// LS Electric XG5000 project: elb
// PLC LSPLC
// module base 0 slot 0: 입출력 모듈:XBC-DR32H (DC 24V 입력, 릴레이 출력 32점)
// module base 0 slot 1: 입력 모듈:XBE-DC16A/B (DC24V 입력, 16점 / DC12/24V 입력, 16점)

PROGRAM 스위치_입력 (task: 스캔 프로그램)

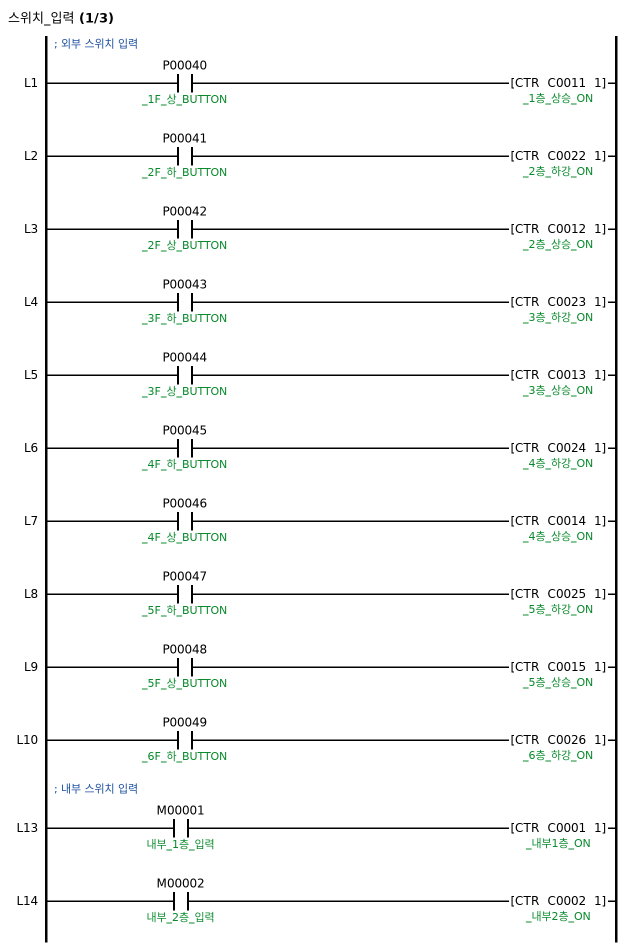
// 외부 스위치 입력
; L1
LOAD      P00040	// _1F_상_BUTTON
CTR       C0011 1	// _1층_상승_ON
; L2
LOAD      P00041	// _2F_하_BUTTON
CTR       C0022 1	// _2층_하강_ON
; L3
LOAD      P00042	// _2F_상_BUTTON
CTR       C0012 1	// _2층_상승_ON
; L4
LOAD      P00043	// _3F_하_BUTTON
CTR       C0023 1	// _3층_하강_ON
; L5
LOAD      P00044	// _3F_상_BUTTON
CTR       C0013 1	// _3층_상승_ON
; L6
LOAD      P00045	// _4F_하_BUTTON
CTR       C0024 1	// _4층_하강_ON
; L7
LOAD      P00046	// _4F_상_BUTTON
CTR       C0014 1	// _4층_상승_ON
; L8
LOAD      P00047	// _5F_하_BUTTON
CTR       C0025 1	// _5층_하강_ON
; L9
LOAD      P00048	// _5F_상_BUTTON
CTR       C0015 1	// _5층_상승_ON
; L10
LOAD      P00049	// _6F_하_BUTTON
CTR       C0026 1	// _6층_하강_ON
// 내부 스위치 입력
; L13
LOAD      M00001	// 내부_1층_입력
CTR       C0001 1	// _내부1층_ON
; L14
LOAD      M00002	// 내부_2층_입력
CTR       C0002 1	// _내부2층_ON

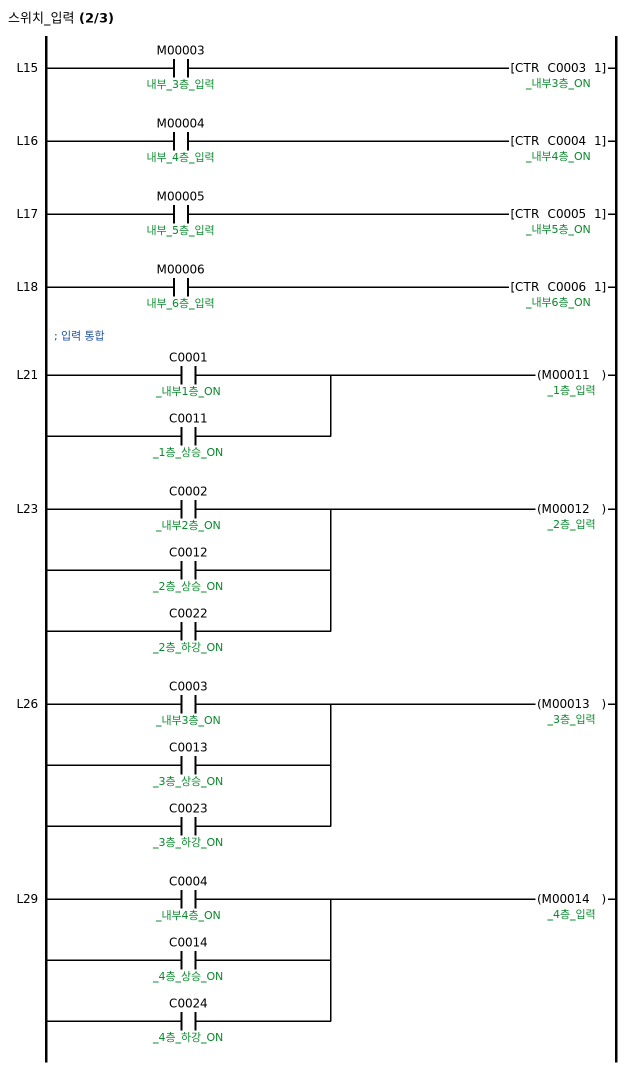
; L15
LOAD      M00003	// 내부_3층_입력
CTR       C0003 1	// _내부3층_ON
; L16
LOAD      M00004	// 내부_4층_입력
CTR       C0004 1	// _내부4층_ON
; L17
LOAD      M00005	// 내부_5층_입력
CTR       C0005 1	// _내부5층_ON
; L18
LOAD      M00006	// 내부_6층_입력
CTR       C0006 1	// _내부6층_ON
// 입력 통합
; L21
LOAD      C0001	// _내부1층_ON
OR        C0011	// _1층_상승_ON
OUT       M00011	// _1층_입력
; L23
LOAD      C0002	// _내부2층_ON
OR        C0012	// _2층_상승_ON
OR        C0022	// _2층_하강_ON
OUT       M00012	// _2층_입력
; L26
LOAD      C0003	// _내부3층_ON
OR        C0013	// _3층_상승_ON
OR        C0023	// _3층_하강_ON
OUT       M00013	// _3층_입력
; L29
LOAD      C0004	// _내부4층_ON
OR        C0014	// _4층_상승_ON
OR        C0024	// _4층_하강_ON
OUT       M00014	// _4층_입력

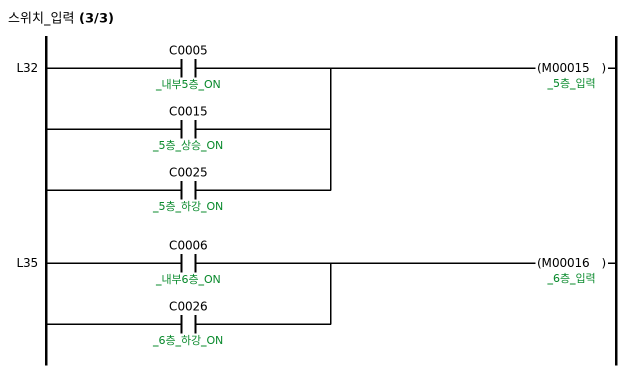
; L32
LOAD      C0005	// _내부5층_ON
OR        C0015	// _5층_상승_ON
OR        C0025	// _5층_하강_ON
OUT       M00015	// _5층_입력
; L35
LOAD      C0006	// _내부6층_ON
OR        C0026	// _6층_하강_ON
OUT       M00016	// _6층_입력

PROGRAM 센서감지(현재위치 (task: 스캔 프로그램)

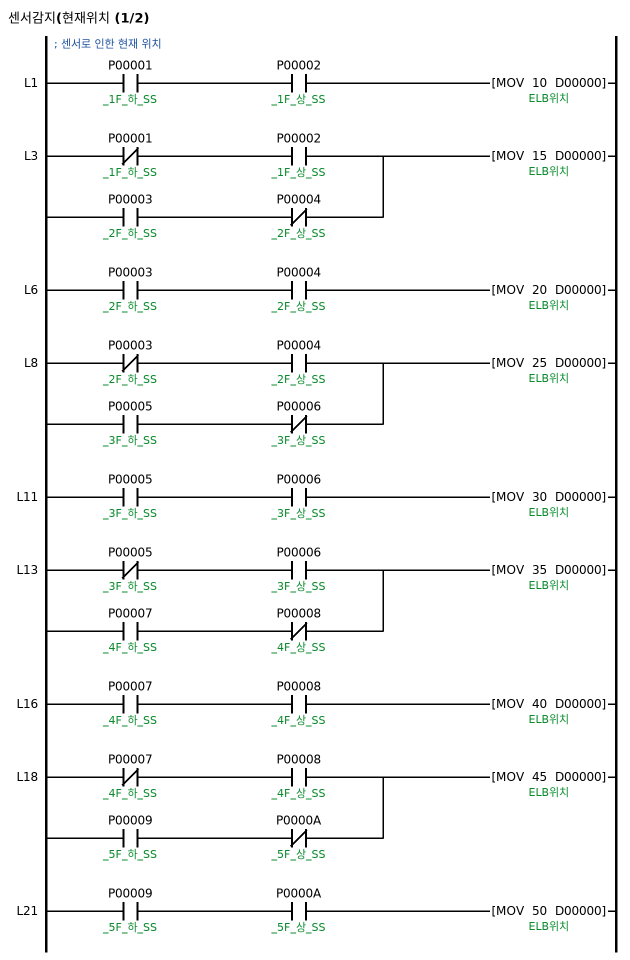
// 센서로 인한 현재 위치
; L1
LOAD      P00001	// _1F_하_SS
AND       P00002	// _1F_상_SS
MOV       10 D00000	// ELB위치
; L3
LOAD NOT  P00001	// _1F_하_SS
AND       P00002	// _1F_상_SS
LOAD      P00003	// _2F_하_SS
AND NOT   P00004	// _2F_상_SS
OR LOAD
MOV       15 D00000	// ELB위치
; L6
LOAD      P00003	// _2F_하_SS
AND       P00004	// _2F_상_SS
MOV       20 D00000	// ELB위치
; L8
LOAD NOT  P00003	// _2F_하_SS
AND       P00004	// _2F_상_SS
LOAD      P00005	// _3F_하_SS
AND NOT   P00006	// _3F_상_SS
OR LOAD
MOV       25 D00000	// ELB위치
; L11
LOAD      P00005	// _3F_하_SS
AND       P00006	// _3F_상_SS
MOV       30 D00000	// ELB위치
; L13
LOAD NOT  P00005	// _3F_하_SS
AND       P00006	// _3F_상_SS
LOAD      P00007	// _4F_하_SS
AND NOT   P00008	// _4F_상_SS
OR LOAD
MOV       35 D00000	// ELB위치
; L16
LOAD      P00007	// _4F_하_SS
AND       P00008	// _4F_상_SS
MOV       40 D00000	// ELB위치
; L18
LOAD NOT  P00007	// _4F_하_SS
AND       P00008	// _4F_상_SS
LOAD      P00009	// _5F_하_SS
AND NOT   P0000A	// _5F_상_SS
OR LOAD
MOV       45 D00000	// ELB위치
; L21
LOAD      P00009	// _5F_하_SS
AND       P0000A	// _5F_상_SS
MOV       50 D00000	// ELB위치

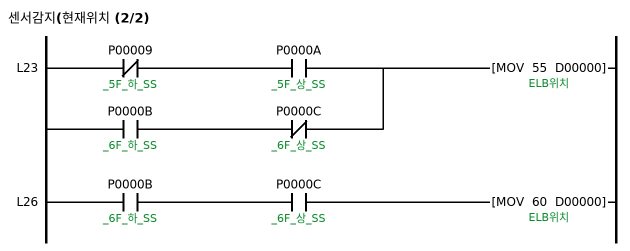
; L23
LOAD NOT  P00009	// _5F_하_SS
AND       P0000A	// _5F_상_SS
LOAD      P0000B	// _6F_하_SS
AND NOT   P0000C	// _6F_상_SS
OR LOAD
MOV       55 D00000	// ELB위치
; L26
LOAD      P0000B	// _6F_하_SS
AND       P0000C	// _6F_상_SS
MOV       60 D00000	// ELB위치

PROGRAM 모드전환 (task: 스캔 프로그램)

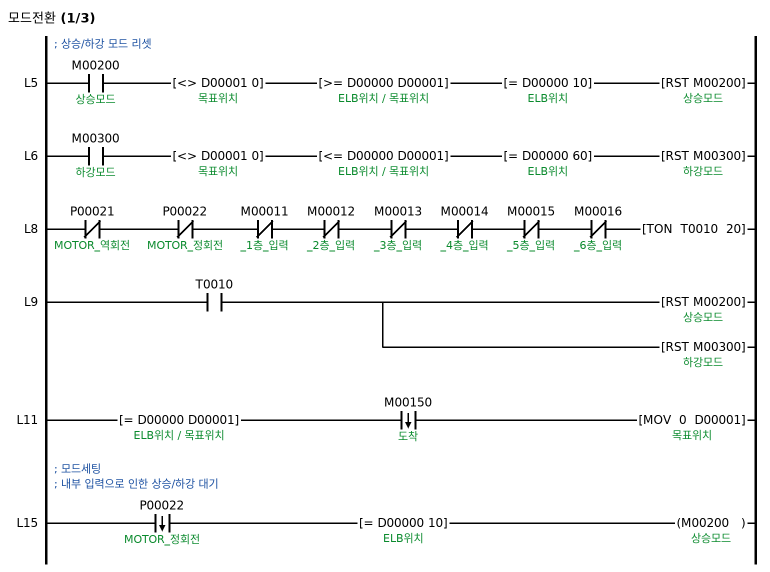
// 상승/하강 모드 리셋
; L5
LOAD      M00200	// 상승모드
AND<>     D00001 0	// 목표위치
AND>=     D00000 D00001	// ELB위치 / 목표위치
AND=      D00000 10	// ELB위치
RST       M00200	// 상승모드
; L6
LOAD      M00300	// 하강모드
AND<>     D00001 0	// 목표위치
AND<=     D00000 D00001	// ELB위치 / 목표위치
AND=      D00000 60	// ELB위치
RST       M00300	// 하강모드
; L8
LOAD NOT  P00021	// MOTOR_역회전
AND NOT   P00022	// MOTOR_정회전
AND NOT   M00011	// _1층_입력
AND NOT   M00012	// _2층_입력
AND NOT   M00013	// _3층_입력
AND NOT   M00014	// _4층_입력
AND NOT   M00015	// _5층_입력
AND NOT   M00016	// _6층_입력
TON       T0010 20
; L9
LOAD      T0010
RST       M00200	// 상승모드
RST       M00300	// 하강모드
; L11
LOAD=     D00000 D00001	// ELB위치 / 목표위치
ANDN      M00150	// 도착
MOV       0 D00001	// 목표위치
// 모드세팅
// 내부 입력으로 인한 상승/하강 대기
; L15
LOADN     P00022	// MOTOR_정회전
AND=      D00000 10	// ELB위치
OUT       M00200	// 상승모드

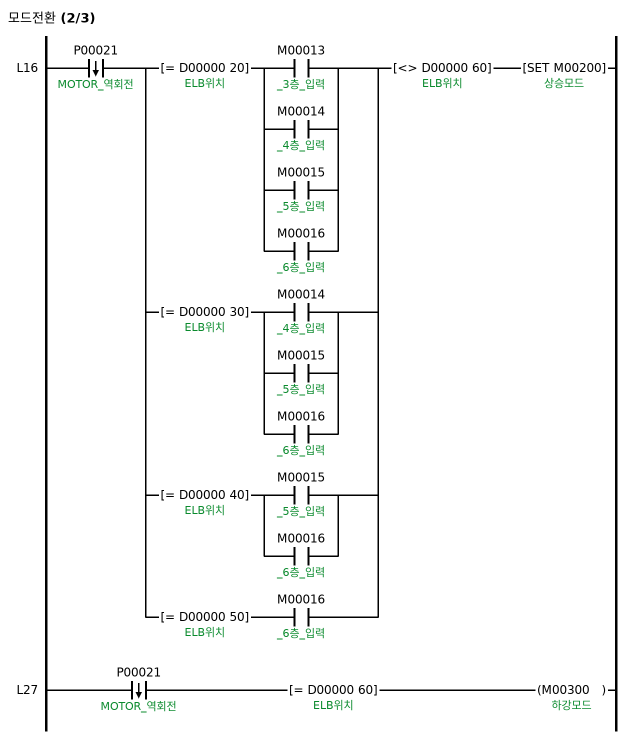
; L16
LOADN     P00021	// MOTOR_역회전
LOAD=     D00000 20	// ELB위치
LOAD      M00013	// _3층_입력
OR        M00014	// _4층_입력
OR        M00015	// _5층_입력
OR        M00016	// _6층_입력
AND LOAD
LOAD=     D00000 30	// ELB위치
LOAD      M00014	// _4층_입력
OR        M00015	// _5층_입력
OR        M00016	// _6층_입력
AND LOAD
OR LOAD
LOAD=     D00000 40	// ELB위치
LOAD      M00015	// _5층_입력
OR        M00016	// _6층_입력
AND LOAD
OR LOAD
LOAD=     D00000 50	// ELB위치
AND       M00016	// _6층_입력
OR LOAD
AND LOAD
AND<>     D00000 60	// ELB위치
SET       M00200	// 상승모드
; L27
LOADN     P00021	// MOTOR_역회전
AND=      D00000 60	// ELB위치
OUT       M00300	// 하강모드

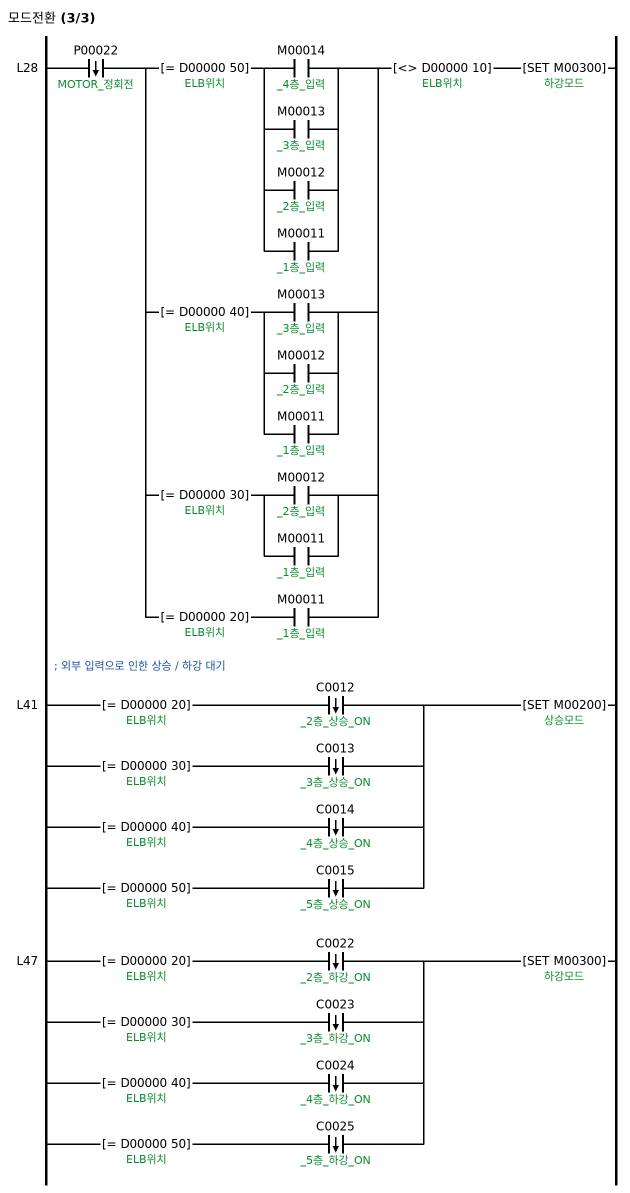
; L28
LOADN     P00022	// MOTOR_정회전
LOAD=     D00000 50	// ELB위치
LOAD      M00014	// _4층_입력
OR        M00013	// _3층_입력
OR        M00012	// _2층_입력
OR        M00011	// _1층_입력
AND LOAD
LOAD=     D00000 40	// ELB위치
LOAD      M00013	// _3층_입력
OR        M00012	// _2층_입력
OR        M00011	// _1층_입력
AND LOAD
OR LOAD
LOAD=     D00000 30	// ELB위치
LOAD      M00012	// _2층_입력
OR        M00011	// _1층_입력
AND LOAD
OR LOAD
LOAD=     D00000 20	// ELB위치
AND       M00011	// _1층_입력
OR LOAD
AND LOAD
AND<>     D00000 10	// ELB위치
SET       M00300	// 하강모드
// 외부 입력으로 인한 상승 / 하강 대기
; L41
LOAD=     D00000 20	// ELB위치
ANDN      C0012	// _2층_상승_ON
LOAD=     D00000 30	// ELB위치
ANDN      C0013	// _3층_상승_ON
OR LOAD
LOAD=     D00000 40	// ELB위치
ANDN      C0014	// _4층_상승_ON
OR LOAD
LOAD=     D00000 50	// ELB위치
ANDN      C0015	// _5층_상승_ON
OR LOAD
SET       M00200	// 상승모드
; L47
LOAD=     D00000 20	// ELB위치
ANDN      C0022	// _2층_하강_ON
LOAD=     D00000 30	// ELB위치
ANDN      C0023	// _3층_하강_ON
OR LOAD
LOAD=     D00000 40	// ELB위치
ANDN      C0024	// _4층_하강_ON
OR LOAD
LOAD=     D00000 50	// ELB위치
ANDN      C0025	// _5층_하강_ON
OR LOAD
SET       M00300	// 하강모드

PROGRAM 스위치리셋 (task: 스캔 프로그램)

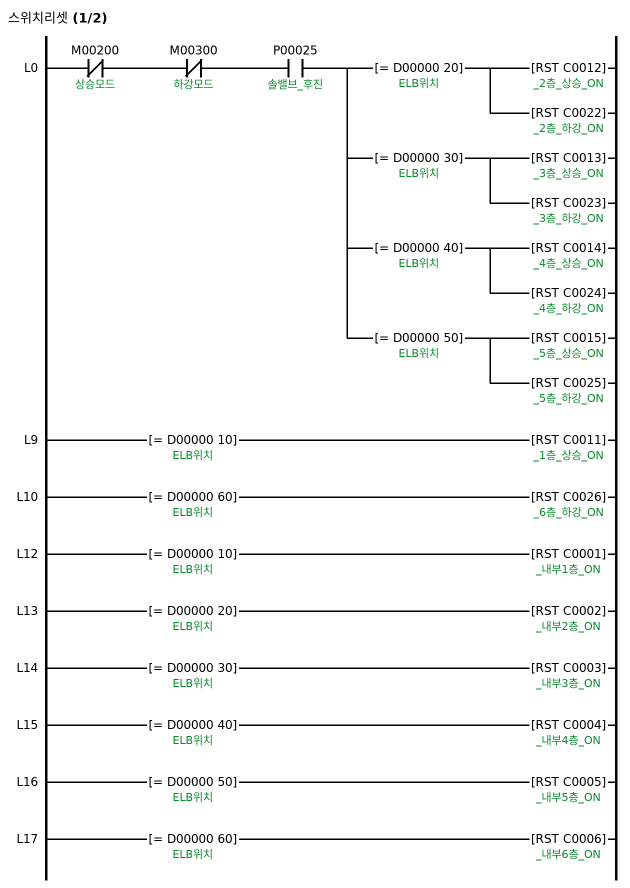
; L0
LOAD NOT  M00200	// 상승모드
AND NOT   M00300	// 하강모드
AND       P00025	// 솔밸브_후진
MPUSH
AND=      D00000 20	// ELB위치
RST       C0012	// _2층_상승_ON
RST       C0022	// _2층_하강_ON
MLOAD
AND=      D00000 30	// ELB위치
RST       C0013	// _3층_상승_ON
RST       C0023	// _3층_하강_ON
MLOAD
AND=      D00000 40	// ELB위치
RST       C0014	// _4층_상승_ON
RST       C0024	// _4층_하강_ON
MPOP
AND=      D00000 50	// ELB위치
RST       C0015	// _5층_상승_ON
RST       C0025	// _5층_하강_ON
; L9
LOAD=     D00000 10	// ELB위치
RST       C0011	// _1층_상승_ON
; L10
LOAD=     D00000 60	// ELB위치
RST       C0026	// _6층_하강_ON
; L12
LOAD=     D00000 10	// ELB위치
RST       C0001	// _내부1층_ON
; L13
LOAD=     D00000 20	// ELB위치
RST       C0002	// _내부2층_ON
; L14
LOAD=     D00000 30	// ELB위치
RST       C0003	// _내부3층_ON
; L15
LOAD=     D00000 40	// ELB위치
RST       C0004	// _내부4층_ON
; L16
LOAD=     D00000 50	// ELB위치
RST       C0005	// _내부5층_ON
; L17
LOAD=     D00000 60	// ELB위치
RST       C0006	// _내부6층_ON

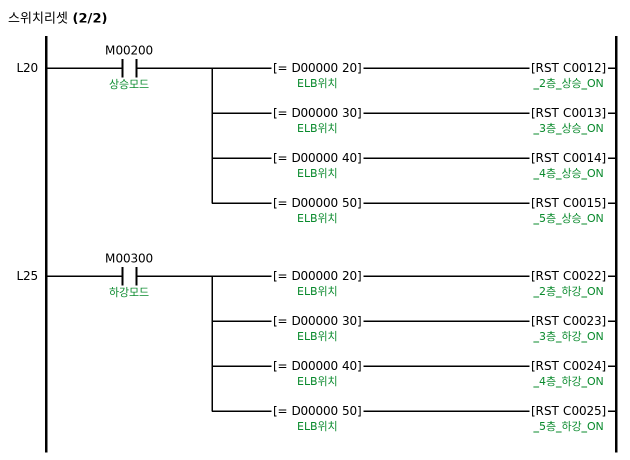
; L20
LOAD      M00200	// 상승모드
MPUSH
AND=      D00000 20	// ELB위치
RST       C0012	// _2층_상승_ON
MLOAD
AND=      D00000 30	// ELB위치
RST       C0013	// _3층_상승_ON
MLOAD
AND=      D00000 40	// ELB위치
RST       C0014	// _4층_상승_ON
MPOP
AND=      D00000 50	// ELB위치
RST       C0015	// _5층_상승_ON
; L25
LOAD      M00300	// 하강모드
MPUSH
AND=      D00000 20	// ELB위치
RST       C0022	// _2층_하강_ON
MLOAD
AND=      D00000 30	// ELB위치
RST       C0023	// _3층_하강_ON
MLOAD
AND=      D00000 40	// ELB위치
RST       C0024	// _4층_하강_ON
MPOP
AND=      D00000 50	// ELB위치
RST       C0025	// _5층_하강_ON

PROGRAM 층수입력 (task: 스캔 프로그램)

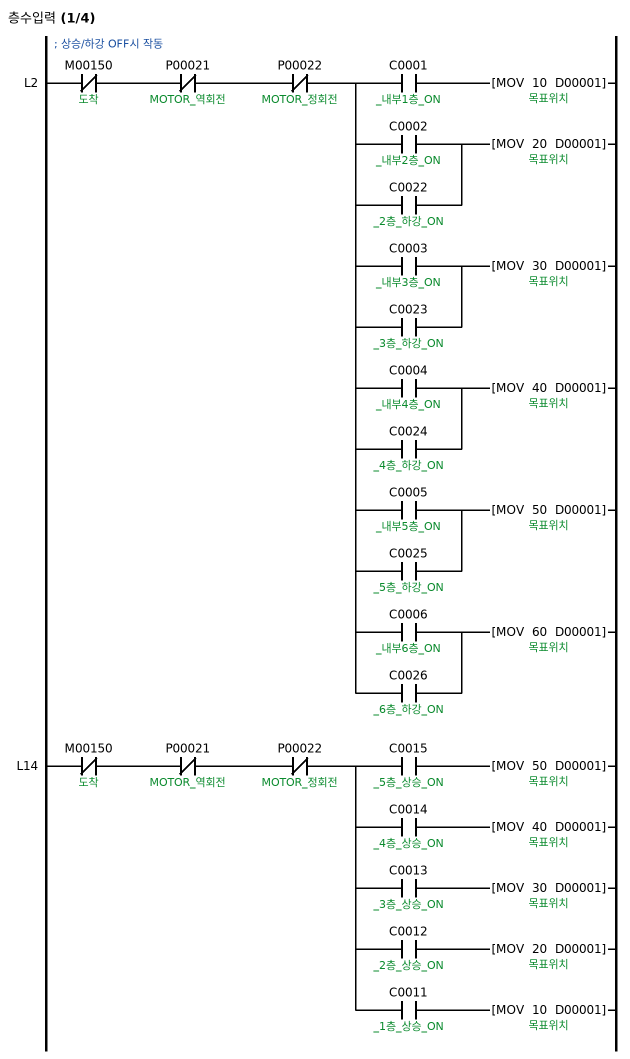
// 상승/하강 OFF시 작동
; L2
LOAD NOT  M00150	// 도착
AND NOT   P00021	// MOTOR_역회전
AND NOT   P00022	// MOTOR_정회전
MPUSH
AND       C0001	// _내부1층_ON
MOV       10 D00001	// 목표위치
MLOAD
LOAD      C0002	// _내부2층_ON
OR        C0022	// _2층_하강_ON
AND LOAD
MOV       20 D00001	// 목표위치
MLOAD
LOAD      C0003	// _내부3층_ON
OR        C0023	// _3층_하강_ON
AND LOAD
MOV       30 D00001	// 목표위치
MLOAD
LOAD      C0004	// _내부4층_ON
OR        C0024	// _4층_하강_ON
AND LOAD
MOV       40 D00001	// 목표위치
MLOAD
LOAD      C0005	// _내부5층_ON
OR        C0025	// _5층_하강_ON
AND LOAD
MOV       50 D00001	// 목표위치
MPOP
LOAD      C0006	// _내부6층_ON
OR        C0026	// _6층_하강_ON
AND LOAD
MOV       60 D00001	// 목표위치
; L14
LOAD NOT  M00150	// 도착
AND NOT   P00021	// MOTOR_역회전
AND NOT   P00022	// MOTOR_정회전
MPUSH
AND       C0015	// _5층_상승_ON
MOV       50 D00001	// 목표위치
MLOAD
AND       C0014	// _4층_상승_ON
MOV       40 D00001	// 목표위치
MLOAD
AND       C0013	// _3층_상승_ON
MOV       30 D00001	// 목표위치
MLOAD
AND       C0012	// _2층_상승_ON
MOV       20 D00001	// 목표위치
MPOP
AND       C0011	// _1층_상승_ON
MOV       10 D00001	// 목표위치

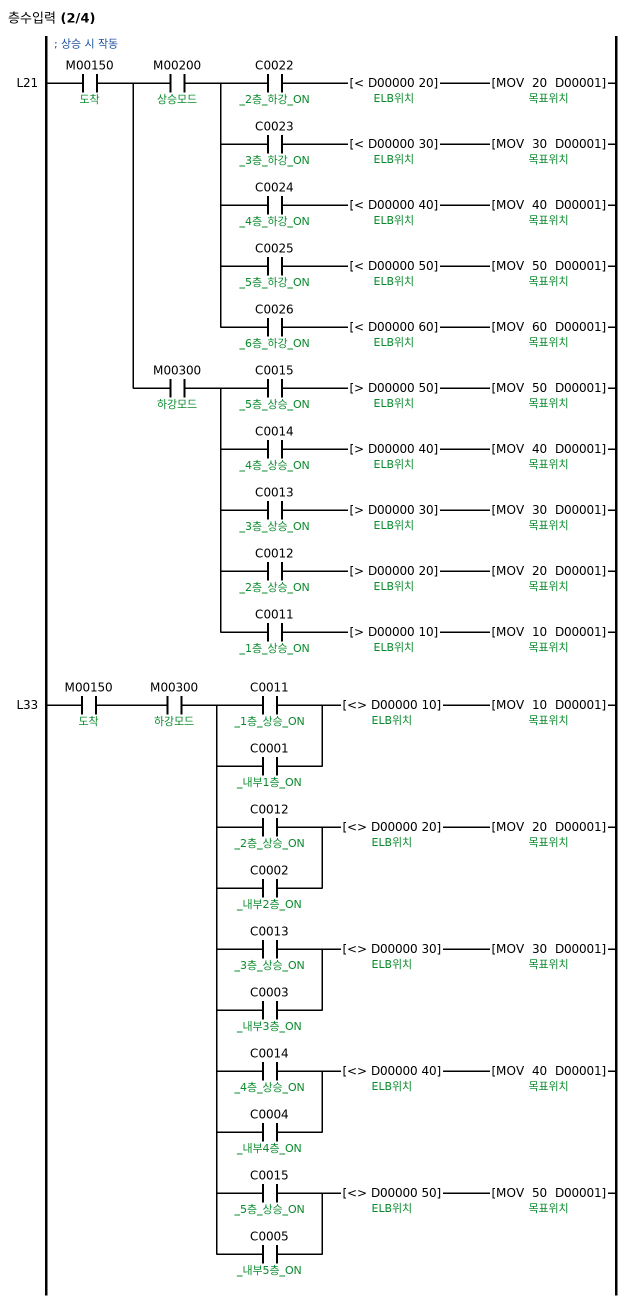
// 상승 시 작동
; L21
LOAD      M00150	// 도착
MPUSH
AND       M00200	// 상승모드
MPUSH
AND       C0022	// _2층_하강_ON
AND<      D00000 20	// ELB위치
MOV       20 D00001	// 목표위치
MLOAD
AND       C0023	// _3층_하강_ON
AND<      D00000 30	// ELB위치
MOV       30 D00001	// 목표위치
MLOAD
AND       C0024	// _4층_하강_ON
AND<      D00000 40	// ELB위치
MOV       40 D00001	// 목표위치
MLOAD
AND       C0025	// _5층_하강_ON
AND<      D00000 50	// ELB위치
MOV       50 D00001	// 목표위치
MPOP
AND       C0026	// _6층_하강_ON
AND<      D00000 60	// ELB위치
MOV       60 D00001	// 목표위치
MPOP
AND       M00300	// 하강모드
MPUSH
AND       C0015	// _5층_상승_ON
AND>      D00000 50	// ELB위치
MOV       50 D00001	// 목표위치
MLOAD
AND       C0014	// _4층_상승_ON
AND>      D00000 40	// ELB위치
MOV       40 D00001	// 목표위치
MLOAD
AND       C0013	// _3층_상승_ON
AND>      D00000 30	// ELB위치
MOV       30 D00001	// 목표위치
MLOAD
AND       C0012	// _2층_상승_ON
AND>      D00000 20	// ELB위치
MOV       20 D00001	// 목표위치
MPOP
AND       C0011	// _1층_상승_ON
AND>      D00000 10	// ELB위치
MOV       10 D00001	// 목표위치
; L33
LOAD      M00150	// 도착
AND       M00300	// 하강모드
MPUSH
LOAD      C0011	// _1층_상승_ON
OR        C0001	// _내부1층_ON
AND LOAD
AND<>     D00000 10	// ELB위치
MOV       10 D00001	// 목표위치
MLOAD
LOAD      C0012	// _2층_상승_ON
OR        C0002	// _내부2층_ON
AND LOAD
AND<>     D00000 20	// ELB위치
MOV       20 D00001	// 목표위치
MLOAD
LOAD      C0013	// _3층_상승_ON
OR        C0003	// _내부3층_ON
AND LOAD
AND<>     D00000 30	// ELB위치
MOV       30 D00001	// 목표위치
MLOAD
LOAD      C0014	// _4층_상승_ON
OR        C0004	// _내부4층_ON
AND LOAD
AND<>     D00000 40	// ELB위치
MOV       40 D00001	// 목표위치
MPOP
LOAD      C0015	// _5층_상승_ON
OR        C0005	// _내부5층_ON
AND LOAD
AND<>     D00000 50	// ELB위치
MOV       50 D00001	// 목표위치

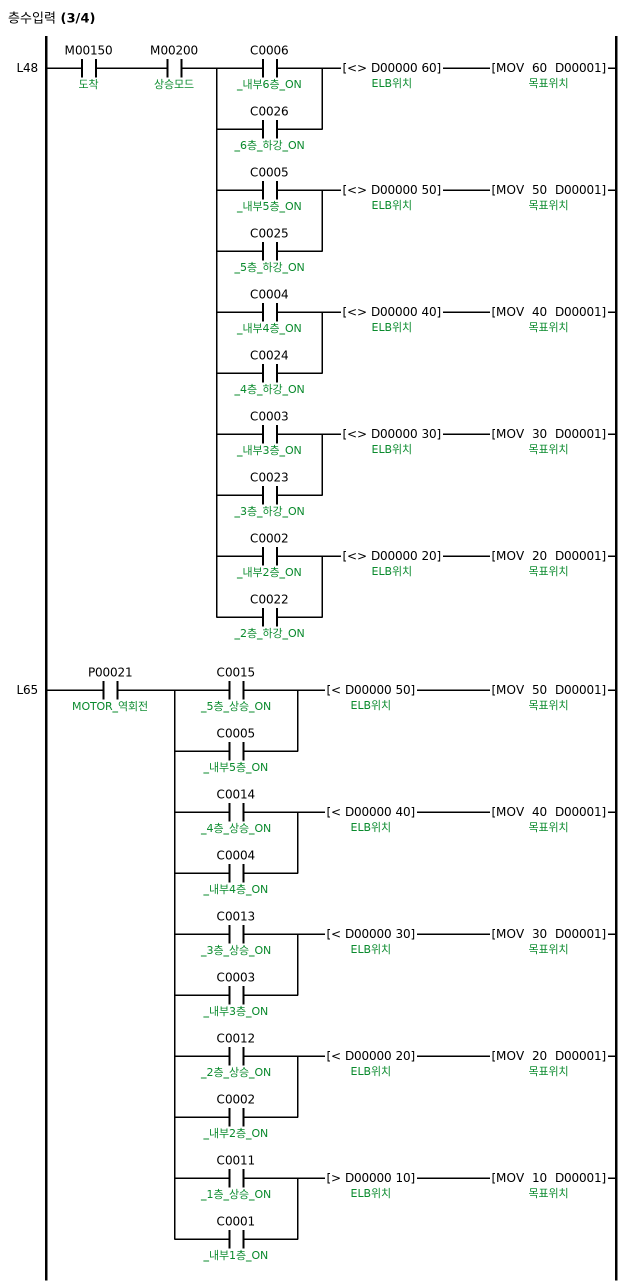
; L48
LOAD      M00150	// 도착
AND       M00200	// 상승모드
MPUSH
LOAD      C0006	// _내부6층_ON
OR        C0026	// _6층_하강_ON
AND LOAD
AND<>     D00000 60	// ELB위치
MOV       60 D00001	// 목표위치
MLOAD
LOAD      C0005	// _내부5층_ON
OR        C0025	// _5층_하강_ON
AND LOAD
AND<>     D00000 50	// ELB위치
MOV       50 D00001	// 목표위치
MLOAD
LOAD      C0004	// _내부4층_ON
OR        C0024	// _4층_하강_ON
AND LOAD
AND<>     D00000 40	// ELB위치
MOV       40 D00001	// 목표위치
MLOAD
LOAD      C0003	// _내부3층_ON
OR        C0023	// _3층_하강_ON
AND LOAD
AND<>     D00000 30	// ELB위치
MOV       30 D00001	// 목표위치
MPOP
LOAD      C0002	// _내부2층_ON
OR        C0022	// _2층_하강_ON
AND LOAD
AND<>     D00000 20	// ELB위치
MOV       20 D00001	// 목표위치
; L65
LOAD      P00021	// MOTOR_역회전
MPUSH
LOAD      C0015	// _5층_상승_ON
OR        C0005	// _내부5층_ON
AND LOAD
AND<      D00000 50	// ELB위치
MOV       50 D00001	// 목표위치
MLOAD
LOAD      C0014	// _4층_상승_ON
OR        C0004	// _내부4층_ON
AND LOAD
AND<      D00000 40	// ELB위치
MOV       40 D00001	// 목표위치
MLOAD
LOAD      C0013	// _3층_상승_ON
OR        C0003	// _내부3층_ON
AND LOAD
AND<      D00000 30	// ELB위치
MOV       30 D00001	// 목표위치
MLOAD
LOAD      C0012	// _2층_상승_ON
OR        C0002	// _내부2층_ON
AND LOAD
AND<      D00000 20	// ELB위치
MOV       20 D00001	// 목표위치
MPOP
LOAD      C0011	// _1층_상승_ON
OR        C0001	// _내부1층_ON
AND LOAD
AND>      D00000 10	// ELB위치
MOV       10 D00001	// 목표위치

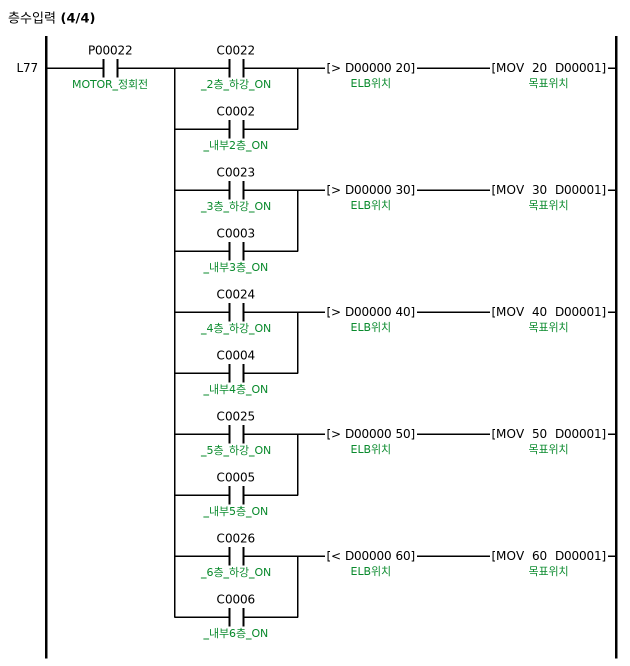
; L77
LOAD      P00022	// MOTOR_정회전
MPUSH
LOAD      C0022	// _2층_하강_ON
OR        C0002	// _내부2층_ON
AND LOAD
AND>      D00000 20	// ELB위치
MOV       20 D00001	// 목표위치
MLOAD
LOAD      C0023	// _3층_하강_ON
OR        C0003	// _내부3층_ON
AND LOAD
AND>      D00000 30	// ELB위치
MOV       30 D00001	// 목표위치
MLOAD
LOAD      C0024	// _4층_하강_ON
OR        C0004	// _내부4층_ON
AND LOAD
AND>      D00000 40	// ELB위치
MOV       40 D00001	// 목표위치
MLOAD
LOAD      C0025	// _5층_하강_ON
OR        C0005	// _내부5층_ON
AND LOAD
AND>      D00000 50	// ELB위치
MOV       50 D00001	// 목표위치
MPOP
LOAD      C0026	// _6층_하강_ON
OR        C0006	// _내부6층_ON
AND LOAD
AND<      D00000 60	// ELB위치
MOV       60 D00001	// 목표위치

PROGRAM 도착 (task: 스캔 프로그램)

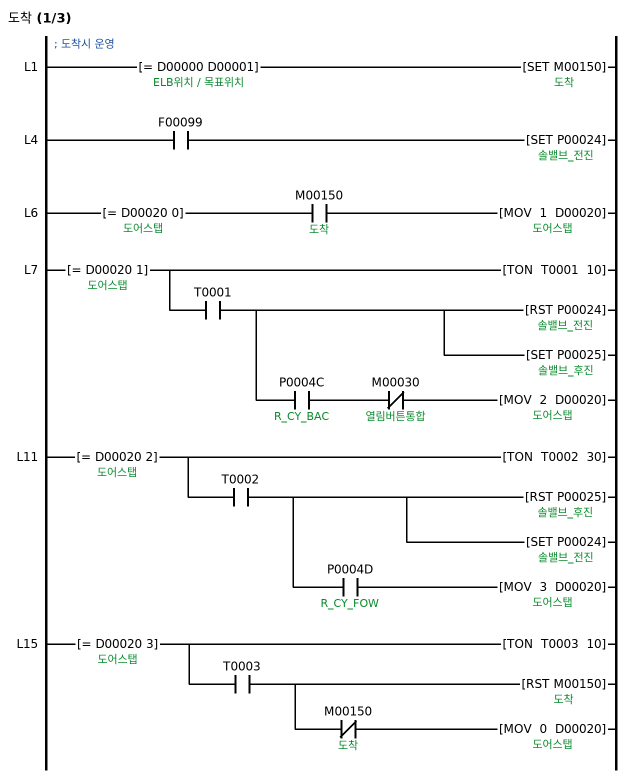
// 도착시 운영
; L1
LOAD=     D00000 D00001	// ELB위치 / 목표위치
SET       M00150	// 도착
; L4
LOAD      F00099
SET       P00024	// 솔밸브_전진
; L6
LOAD=     D00020 0	// 도어스탭
AND       M00150	// 도착
MOV       1 D00020	// 도어스탭
; L7
LOAD=     D00020 1	// 도어스탭
TON       T0001 10
AND       T0001
RST       P00024	// 솔밸브_전진
SET       P00025	// 솔밸브_후진
AND       P0004C	// R_CY_BAC
AND NOT   M00030	// 열림버튼통합
MOV       2 D00020	// 도어스탭
; L11
LOAD=     D00020 2	// 도어스탭
TON       T0002 30
AND       T0002
RST       P00025	// 솔밸브_후진
SET       P00024	// 솔밸브_전진
AND       P0004D	// R_CY_FOW
MOV       3 D00020	// 도어스탭
; L15
LOAD=     D00020 3	// 도어스탭
TON       T0003 10
AND       T0003
RST       M00150	// 도착
AND NOT   M00150	// 도착
MOV       0 D00020	// 도어스탭

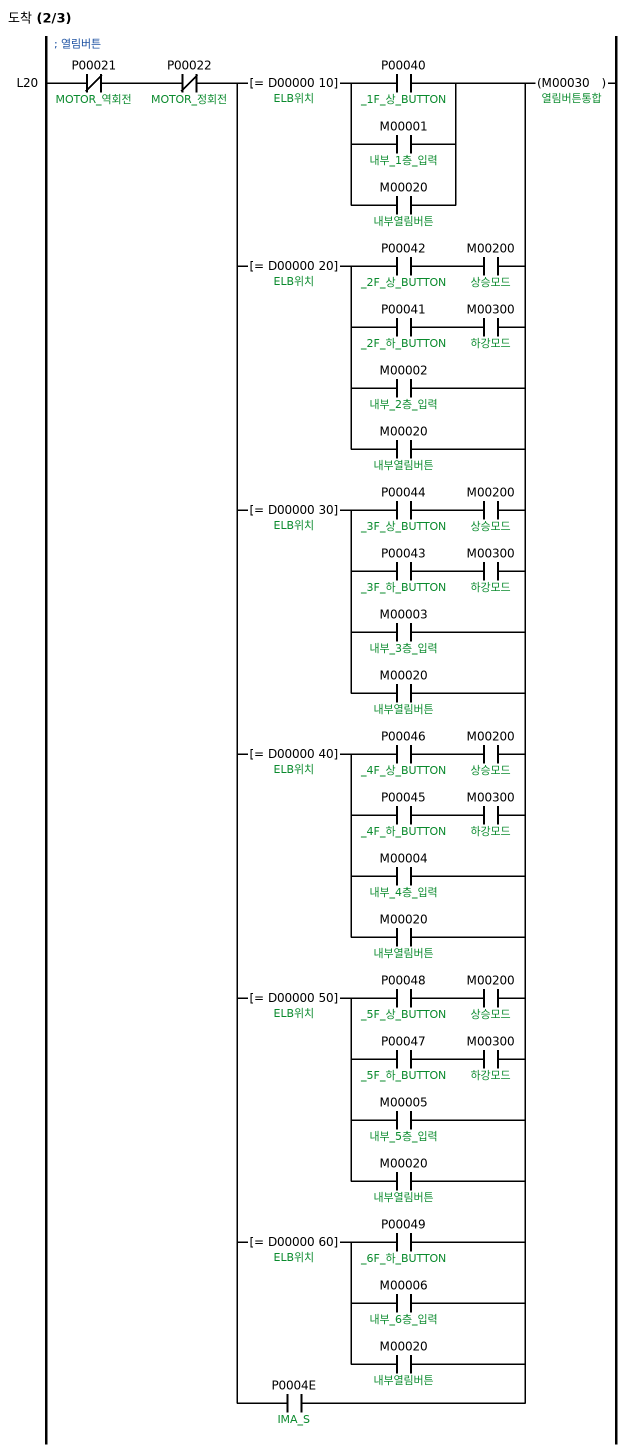
// 열림버튼
; L20
LOAD NOT  P00021	// MOTOR_역회전
AND NOT   P00022	// MOTOR_정회전
LOAD=     D00000 10	// ELB위치
LOAD      P00040	// _1F_상_BUTTON
OR        M00001	// 내부_1층_입력
OR        M00020	// 내부열림버튼
AND LOAD
LOAD=     D00000 20	// ELB위치
LOAD      P00042	// _2F_상_BUTTON
AND       M00200	// 상승모드
LOAD      P00041	// _2F_하_BUTTON
AND       M00300	// 하강모드
OR LOAD
OR        M00002	// 내부_2층_입력
OR        M00020	// 내부열림버튼
AND LOAD
OR LOAD
LOAD=     D00000 30	// ELB위치
LOAD      P00044	// _3F_상_BUTTON
AND       M00200	// 상승모드
LOAD      P00043	// _3F_하_BUTTON
AND       M00300	// 하강모드
OR LOAD
OR        M00003	// 내부_3층_입력
OR        M00020	// 내부열림버튼
AND LOAD
OR LOAD
LOAD=     D00000 40	// ELB위치
LOAD      P00046	// _4F_상_BUTTON
AND       M00200	// 상승모드
LOAD      P00045	// _4F_하_BUTTON
AND       M00300	// 하강모드
OR LOAD
OR        M00004	// 내부_4층_입력
OR        M00020	// 내부열림버튼
AND LOAD
OR LOAD
LOAD=     D00000 50	// ELB위치
LOAD      P00048	// _5F_상_BUTTON
AND       M00200	// 상승모드
LOAD      P00047	// _5F_하_BUTTON
AND       M00300	// 하강모드
OR LOAD
OR        M00005	// 내부_5층_입력
OR        M00020	// 내부열림버튼
AND LOAD
OR LOAD
LOAD=     D00000 60	// ELB위치
LOAD      P00049	// _6F_하_BUTTON
OR        M00006	// 내부_6층_입력
OR        M00020	// 내부열림버튼
AND LOAD
OR LOAD
OR        P0004E	// IMA_S
AND LOAD
OUT       M00030	// 열림버튼통합

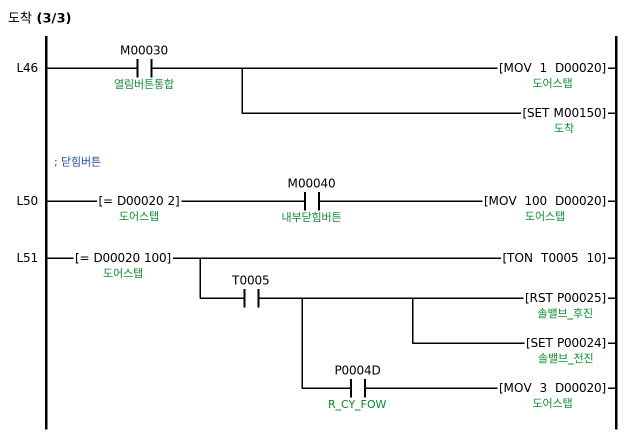
; L46
LOAD      M00030	// 열림버튼통합
MOV       1 D00020	// 도어스탭
SET       M00150	// 도착
// 닫힘버튼
; L50
LOAD=     D00020 2	// 도어스탭
AND       M00040	// 내부닫힘버튼
MOV       100 D00020	// 도어스탭
; L51
LOAD=     D00020 100	// 도어스탭
TON       T0005 10
AND       T0005
RST       P00025	// 솔밸브_후진
SET       P00024	// 솔밸브_전진
AND       P0004D	// R_CY_FOW
MOV       3 D00020	// 도어스탭

PROGRAM 모터구동 (task: 스캔 프로그램)

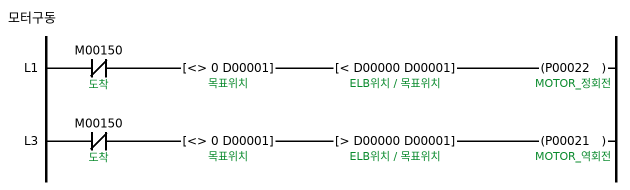
; L1
LOAD NOT  M00150	// 도착
AND<>     0 D00001	// 목표위치
AND<      D00000 D00001	// ELB위치 / 목표위치
OUT       P00022	// MOTOR_정회전
; L3
LOAD NOT  M00150	// 도착
AND<>     0 D00001	// 목표위치
AND>      D00000 D00001	// ELB위치 / 목표위치
OUT       P00021	// MOTOR_역회전

VARIABLES AND COMMENTS (devices not used above)
P0004A	BIT	L_CY_BAC
P0004B	BIT	L_CY_FOW
P0002E	BIT	모터상승
P0004F	BIT	비상정지